// TIA Portal V18 export
FUNCTION "ALARMES" : Void   // FC13, LAD
{ S7_Optimized_Access := 'TRUE' }
// stored: SetENOAutomatically false
BEGIN

REGION Network 1: ALARMES CABINE
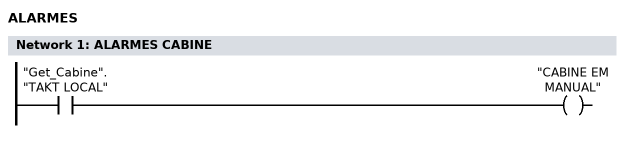
   RUNG wire#powerrail
      Contact( "Get_Cabine"."TAKT LOCAL" )
      Coil( "CABINE EM MANUAL" )
   END_RUNG
   // the same network as SCL:
   "CABINE EM MANUAL" := "Get_Cabine"."TAKT LOCAL";
END_REGION
END_FUNCTION
